Fanuc KAREL source: kc00037.KL

-- PROVISIONAL review KL for V940-1; original PC SHA256 72dd9edeec05af5ab245ad2cf34beef6a580d18ed2ad0ec8c941b8417c6e908f
-- Incomplete behavior may be omitted. Consult companion uncertainty JSON. Do not deploy.
PROGRAM KC00037
%NOLOCKGROUP
BEGIN
  -- V9_ZERO_TABLE_METADATA_HINT layout=0002_ascii; no indexed target words; source/name/runtime held
  -- UNRESOLVED_PC offsets 5-29; opcodes 27,22,2A,22,22,31
  -- UNRESOLVED_PC offsets 34-38; opcodes 7F
END KC00037
